// TIA Portal V19 export
// export: Created 2026-10-15T09:44:25.0145674Z, ExportSetting WithDefaults, DisplayName Totally Integrated Automation Portal, DisplayVersion V19, DisplayName TIA Portal Openness, DisplayVersion V19, DisplayName TIA Portal Version Control Interface, DisplayVersion V19, DisplayName STEP 7 Professional, DisplayVersion V19, DisplayName STEP 7 Safety, DisplayVersion V19, DisplayName WinCC Basic/Comfort/Advanced, DisplayVersion V19, DisplayName WinCC Unified, DisplayVersion V19
FUNCTION "ROLL_PB51" : Void   // FC34, SCL
{ S7_Optimized_Access := 'TRUE' }
VERSION : 0.1
// stored: AutoNumber true, IsIECCheckEnabled false, SetENOAutomatically false, UDAEnableTagReadback false
   VAR_TEMP
      r : Bool;
      a1 : Word;
      a2 : Word;
      activeDataBlock : Int;
      comparisonResults : Array[0..0] of Bool;
   END_VAR
BEGIN

   #r := FALSE;
   #a1 := W#16#0000;
   #a2 := W#16#0000;
   #activeDataBlock := 0;
   // PB51, STEP 5 network 1
   #a2 := #a1;
   #a1 := W#16#2060;
   #r := "ROLL_IO".Output[24, 0];
   "ROLL_TimerOp"(Number := 15,
                  Operation := 0,
                  Signal := #r,
                  Preset := #a1);
   // PB51, STEP 5 network 2
   #a2 := #a1;
   #a1 := W#16#3360;
   #r := ((NOT "ROLL_IO".Input[5, 6]) AND "ROLL_State".M[31, 5]);
   "ROLL_TimerOp"(Number := 16,
                  Operation := 0,
                  Signal := #r,
                  Preset := #a1);
   // PB51, STEP 5 network 3
   #a2 := #a1;
   #a1 := W#16#1010;
   #r := "ROLL_State".M[37, 5];
   "ROLL_TimerOp"(Number := 18,
                  Operation := 0,
                  Signal := #r,
                  Preset := #a1);
   // PB51, STEP 5 network 4
   #a2 := #a1;
   #a1 := W#16#2015;
   #r := (((NOT "ROLL_IO".Input[124, 1]) AND "ROLL_IO".Output[112, 1]) OR ((NOT "ROLL_IO".Input[124, 2]) AND "ROLL_IO".Output[112, 2]));
   "ROLL_TimerOp"(Number := 19,
                  Operation := 0,
                  Signal := #r,
                  Preset := #a1);
   // PB51, STEP 5 network 5
   #a2 := #a1;
   #a1 := W#16#1010;
   #r := (("ROLL_IO".Input[123, 4] OR "ROLL_IO".Input[123, 5]) AND "ROLL_IO".Output[112, 0]);
   "ROLL_TimerOp"(Number := 20,
                  Operation := 0,
                  Signal := #r,
                  Preset := #a1);
   // PB51, STEP 5 network 6
   #a2 := #a1;
   #a1 := W#16#1050;
   #r := "ROLL_IO".Input[123, 4];
   "ROLL_TimerOp"(Number := 21,
                  Operation := 0,
                  Signal := #r,
                  Preset := #a1);
   // PB51, STEP 5 network 7
   #a2 := #a1;
   #a1 := W#16#2005;
   #r := ("ROLL_IO".Input[125, 0] AND "ROLL_IO".Input[125, 1]);
   "ROLL_TimerOp"(Number := 95,
                  Operation := 0,
                  Signal := #r,
                  Preset := #a1);
   // PB51, STEP 5 network 8
   RETURN;
END_FUNCTION
